(* IEC 61131-3 sources: ZPLC/packages/zplc-ide/plant-scenes/belt-to-belt-transfer, 2 files *)

(* ---- reference.st ---- *)
PROGRAM BeltTransfer
VAR_INPUT
    Start    AT %I0.0 : BOOL;
    Waiting  AT %I0.1 : BOOL;
    OutEye   AT %I0.2 : BOOL;
    XMin     AT %I0.3 : BOOL;
    XMax     AT %I0.4 : BOOL;
    YMin     AT %I0.5 : BOOL;
    YMax     AT %I0.6 : BOOL;
    Gripped  AT %I0.7 : BOOL;
END_VAR
VAR_OUTPUT
    RunIn    AT %Q0.0 : BOOL;
    RunOut   AT %Q0.1 : BOOL;
    Emit     AT %Q0.2 : BOOL;
    Hold     AT %Q0.3 : BOOL;
    XPlus    AT %Q0.4 : BOOL;
    XMinus   AT %Q0.5 : BOOL;
    YPlus    AT %Q0.6 : BOOL;
    YMinus   AT %Q0.7 : BOOL;
    Grip     AT %Q1.0 : BOOL;
    Busy     AT %Q1.1 : BOOL;
    Done     AT %Q1.2 : BOOL;
END_VAR
VAR
    Active    : BOOL;
    State     : INT;
    Emitted   : INT;
    Placed    : INT;
    Feed      : BOOL;
    Settle    : TON;
    Rest      : TON;
    OutRise   : R_TRIG;
    Delivered : CTU;
END_VAR

IF Start THEN
    Active := TRUE;
END_IF;

(* the box must stand still at the blade before the clamp comes down; after the release
   it must lie still on the stopped outfeed belt before the belt runs again *)
Settle(IN := Waiting AND State = 2, PT := T#300ms);
Rest(IN := State = 8, PT := T#600ms);
OutRise(CLK := OutEye);
Delivered(CU := OutRise.Q, R := FALSE, PV := 4);

(* one state per move: 0 idle, 2 wait for a box, 3 lower, 4 close, 5 lift, 6 carry,
   7 lower, 8 open and settle, 9 lift, 10 return, 11 finished *)
CASE State OF
    0:
        IF Active THEN
            Feed := TRUE;
            Emitted := 1;
            State := 2;
        END_IF;
    2:
        IF Settle.Q AND YMax AND XMin THEN
            State := 3;
        END_IF;
    3:
        IF YMin THEN
            State := 4;
        END_IF;
    4:
        IF Gripped THEN
            State := 5;
        END_IF;
    5:
        IF YMax THEN
            (* the box has left the blade: bring the next one while this one is carried *)
            IF Emitted < 4 THEN
                Feed := TRUE;
                Emitted := Emitted + 1;
            END_IF;
            State := 6;
        END_IF;
    6:
        IF XMax THEN
            State := 7;
        END_IF;
    7:
        IF YMin THEN
            State := 8;
        END_IF;
    8:
        IF Rest.Q THEN
            Placed := Placed + 1;
            State := 9;
        END_IF;
    9:
        IF YMax THEN
            State := 10;
        END_IF;
    10:
        IF XMin THEN
            IF Placed < 4 THEN
                State := 2;
            ELSE
                State := 11;
            END_IF;
        END_IF;
END_CASE;

RunIn  := Active;
Hold   := Active;
(* the outfeed belt stands still while a box is carried over it, put down and settling *)
RunOut := Active AND NOT (State = 6 OR State = 7 OR State = 8);
Emit   := Feed;
Feed   := FALSE;
Grip   := State >= 4 AND State <= 7;
YPlus  := (State = 2 OR State = 5 OR State = 9) AND NOT YMax;
YMinus := (State = 3 OR State = 7) AND NOT YMin;
XPlus  := State = 6 AND NOT XMax;
XMinus := (State = 2 OR State = 10) AND NOT XMin;
Done   := Delivered.Q;
Busy   := Active AND NOT Delivered.Q;

END_PROGRAM

(* ---- starter.st ---- *)
PROGRAM BeltTransfer
VAR_INPUT
    Start    AT %I0.0 : BOOL;  (* StartButton.pressed: start the transfer *)
    Waiting  AT %I0.1 : BOOL;  (* EyePick.detect: a box waits at the stop blade of the infeed *)
    OutEye   AT %I0.2 : BOOL;  (* EyeOut.detect: a box passes on the outfeed belt *)
    XMin     AT %I0.3 : BOOL;  (* Pick1.xAtMin: the carriage is over the infeed *)
    XMax     AT %I0.4 : BOOL;  (* Pick1.xAtMax: the carriage is over the outfeed *)
    YMin     AT %I0.5 : BOOL;  (* Pick1.yAtMin: the clamp is down *)
    YMax     AT %I0.6 : BOOL;  (* Pick1.yAtMax: the clamp is up *)
    Gripped  AT %I0.7 : BOOL;  (* Pick1.gripped: the clamp holds a box *)
END_VAR
VAR_OUTPUT
    RunIn    AT %Q0.0 : BOOL;  (* Infeed.run: run the infeed belt *)
    RunOut   AT %Q0.1 : BOOL;  (* Outfeed.run: run the outfeed belt *)
    Emit     AT %Q0.2 : BOOL;  (* Source1.emit: put one box on the infeed belt *)
    Hold     AT %Q0.3 : BOOL;  (* Stop1.extend: the blade holds the box while true *)
    XPlus    AT %Q0.4 : BOOL;  (* Pick1.xPlus: move toward the outfeed while true *)
    XMinus   AT %Q0.5 : BOOL;  (* Pick1.xMinus: move toward the infeed while true *)
    YPlus    AT %Q0.6 : BOOL;  (* Pick1.yPlus: lift the clamp while true *)
    YMinus   AT %Q0.7 : BOOL;  (* Pick1.yMinus: lower the clamp while true *)
    Grip     AT %Q1.0 : BOOL;  (* Pick1.grip: close the clamp while true *)
    Busy     AT %Q1.1 : BOOL;  (* Beacon.amber: the transfer is running *)
    Done     AT %Q1.2 : BOOL;  (* Beacon.green: lit when four boxes have crossed the outfeed *)
END_VAR

(* Goal: a press of the start button runs the infeed and puts four boxes on
   it, one at a time. The blade stops each box where the clamp can reach it.
   For every box: lower the clamp, close it and wait for Gripped, lift, carry
   the box over the outfeed, lower, open the clamp and let the box settle,
   lift, and return. Keep the outfeed belt stopped while a box is put down on
   it and run it afterwards. Light Busy while the transfer runs and Done when
   four boxes have passed EyeOut. *)

END_PROGRAM
